Fanuc KAREL source: CA0110.KL

PROGRAM CA0110
%STACKSIZE=65535
%PRIORITY=65535
%NOLOCKGROUP
TYPE
T=STRUCTURE
A : INTEGER
B : REAL
ENDSTRUCTURE
VAR
G : INTEGER
I : INTEGER
R : REAL
B : BOOLEAN
S : STRING[16]
AI : ARRAY[2] OF INTEGER
AR : ARRAY[2] OF REAL
ST : T
P : XYZWPR
V : VECTOR
ROUTINE F(P1 : BOOLEAN) : BOOLEAN FROM CA0110
ROUTINE F
BEGIN
RETURN(P1)
-- UNRESOLVED_PC line 22 opcodes [7F] marker_code=16
END F
BEGIN
G=0
I=1
R=2.5
B=TRUE
S='A'
AI[1]=3
AR[1]=4.5
-- UNSAFE_SOURCE_IR line 31: ST.A = 5
-- UNSAFE_SOURCE_IR line 32: ST.B = 6.5
-- UNSAFE_SOURCE_IR line 33: CALL_RESULT F(B)
G=(G + 1)
END CA0110
